(* IEC 61131-3 sources: Codesys_IAP/Demo/PLC1/PLC 1 Simulatie Ladder StructuredTekst IOStructures 2V0_tekst/Programma Structured Text/States, 5 files *)

(* ---- magazijnStates.st ---- *)
(*#### DECLARATIE ####*)
// Datum : 17 december 2020, Auteur: Gerard Harkema
{attribute 'qualified_only'}
{attribute 'strict'}
TYPE magazijnStates :
(
	idle := 0,
	in,
	travel_out,
	out,
	travel_in,
	error
);
END_TYPE

(* ---- overzetterStates.st ---- *)
(*#### DECLARATIE ####*)
// Datum : 17 december 2020, Auteur: Gerard Harkema
{attribute 'qualified_only'}
{attribute 'strict'}
TYPE overzetterStates :
(
	idle := 0,
	is_links,
	vaccuum_aanzetten,
	ga_naar_rechts,
	is_rechts,
	vaccuum_lossen,
	ga_naar_midden,
	is_midden,
	ga_naar_links,
	error
);
END_TYPE

(* ---- sorteerStates.st ---- *)
(*#### DECLARATIE ####*)
// Datum : 17 december 2020, Auteur: Gerard Harkema
{attribute 'qualified_only'}
{attribute 'strict'}
TYPE sorteerStates :
(
	idle := 0,
	wacht_op_start,
	stopper_uit,
	meten,
	uitvoer_goot_uit,
	transporteren_naar_goot,
	uitvoer_goot_in,
	goot_vol,
	error,
	reset_error
);
END_TYPE

(* ---- sorteerStationStates.st ---- *)
(*#### DECLARATIE ####*)
// Datum : 17 december 2020, Auteur: Gerard Harkema
{attribute 'qualified_only'}
{attribute 'strict'}
TYPE sorteerStationStates :
(
	idle := 0,
	wacht_op_klaar,
	wacht_enable,
	product_uitgifte,
	product_overzetten,
	product_sorteren,
	service,
	error
);
END_TYPE

(* ---- uitvoerGootStates.st ---- *)
(*#### DECLARATIE ####*)
// Datum : 17 december 2020, Auteur: Gerard Harkema
{attribute 'qualified_only'}
{attribute 'strict'}
TYPE uitvoerGootStates :
(
	idle := 0,
	is_in,
	ga_in,
	is_uit,
	ga_uit,
	error
);
END_TYPE
